FUNCTION StationParameter_28000_1  : BOOL
VAR
  nStationParameter                 : UINT; // THIS IS ONLY FOR EXAMPLE USE, CHECK MAX_STATION MANUALLY
END_VAR

//-----------------------------------------------------------------------------------------------------------------------------------------
//-----------------------------------------------------------------------------------------------------------------------------------------
//
//  HAUD 2026.11.02
//
//  - hard coded station parameters
//  - TODO: xml DataServer implementation for station parameter read/write
//
//  - reminder: (this you HAVE to check manually when setting up the transport)
//-----------------------------------------------------------------------------
//    - DO NOT place the modulo turn within the range of a station
//
//    - in case the extern process requires multiple xts stations, 
//      - the range must be closed and in strict order
//-----------------------------------------------------------------------------------------------------------------------------------------
//-----------------------------------------------------------------------------------------------------------------------------------------
GVL_XTS.StationStartIndex                                         := 142;
GVL_XTS.StationStart.rPosWait                                     :=    5000.0; // for every TRANSPORT_START this physical position may differ from the rPosWait of StationStartIndex station

GVL_XTS.StationStart.rGap                                         :=     110.0;
GVL_XTS.StationStart.rVelo                                        :=   1_250.0;
GVL_XTS.StationStart.rAccDec                                      :=  12_500.0;
GVL_XTS.StationStart.rJerk                                        := 100_000.0;

FOR nStationParameter := 1 TO GVL_XTS_CONSTANTS.MAX_STATION
DO
  GVL_XTS.StationParameter[nStationParameter].eType               := E_STATION_TYPE.STATION_PROCESS;
  GVL_XTS.StationParameter[nStationParameter].rGap                := MAIN_APP.rDefaultGap;
  GVL_XTS.StationParameter[nStationParameter].rVelo               := MAIN_APP.rDefaultVeloMin;
  GVL_XTS.StationParameter[nStationParameter].rAccDec             := MAIN_APP.rDefaultAccDec;
  GVL_XTS.StationParameter[nStationParameter].rJerk               := MAIN_APP.rDefaultJerk;
END_FOR
//-----------------------------------------------------------------------------------------------------------------------------------------
//  PRC 01 reserve
//-----------------------------------------------------------------------------------------------------------------------------------------
FOR nStationParameter := 1 TO 16
DO
  GVL_XTS.StationParameter[nStationParameter].rVelo               := MAIN_APP.rDefaultVeloMin;
END_FOR
nStationParameter := 1;
GVL_XTS.StationParameter[nStationParameter].eType                 := E_STATION_TYPE.STATION_PROCESS;
GVL_XTS.StationParameter[nStationParameter].sText                 := 'PRC_01_01';
GVL_XTS.StationParameter[nStationParameter].nConfiguredStopCount  :=       1;   // how many stops the mover has to make in this station

GVL_XTS.StationParameter[nStationParameter].rPosWait              :=   3000.0+80.0; // absolute modulo position
GVL_XTS.StationParameter[nStationParameter].rPosStop[1]           :=       0.0; // relative to rPosWait
GVL_XTS.StationParameter[nStationParameter].rReleaseDistance      :=    2000.0; // relative to Mover.ActPos

nStationParameter := 2;
GVL_XTS.StationParameter[nStationParameter].eType                 := E_STATION_TYPE.STATION_PROCESS;
GVL_XTS.StationParameter[nStationParameter].sText                 := 'PRC_01_02';
GVL_XTS.StationParameter[nStationParameter].nConfiguredStopCount  :=       1;   // how many stops the mover has to make in this station

GVL_XTS.StationParameter[nStationParameter].rPosWait              :=   3000.0+160.0; // absolute modulo position
GVL_XTS.StationParameter[nStationParameter].rPosStop[1]           :=       0.0; // relative to rPosWait
GVL_XTS.StationParameter[nStationParameter].rReleaseDistance      :=    1900.0; // relative to Mover.ActPos

nStationParameter := 3;
GVL_XTS.StationParameter[nStationParameter].eType                 := E_STATION_TYPE.STATION_PROCESS;
GVL_XTS.StationParameter[nStationParameter].sText                 := 'PRC_01_03';
GVL_XTS.StationParameter[nStationParameter].nConfiguredStopCount  :=       1;   // how many stops the mover has to make in this station

GVL_XTS.StationParameter[nStationParameter].rPosWait              :=     3000.0+240.0; // absolute modulo position
GVL_XTS.StationParameter[nStationParameter].rPosStop[1]           :=       0.0; // relative to rPosWait
GVL_XTS.StationParameter[nStationParameter].rReleaseDistance      :=    1120.0; // relative to Mover.ActPos

nStationParameter := 4;
GVL_XTS.StationParameter[nStationParameter].eType                 := E_STATION_TYPE.STATION_PROCESS;
GVL_XTS.StationParameter[nStationParameter].sText                 := 'PRC_01_04';
GVL_XTS.StationParameter[nStationParameter].nConfiguredStopCount  :=       1;   // how many stops the mover has to make in this station

GVL_XTS.StationParameter[nStationParameter].rPosWait              :=     3000.0+320.0; // absolute modulo position
GVL_XTS.StationParameter[nStationParameter].rPosStop[1]           :=       0.0; // relative to rPosWait
GVL_XTS.StationParameter[nStationParameter].rReleaseDistance      :=    1040.0; // relative to Mover.ActPos

nStationParameter := 5;
GVL_XTS.StationParameter[nStationParameter].eType                 := E_STATION_TYPE.STATION_PROCESS;
GVL_XTS.StationParameter[nStationParameter].sText                 := 'PRC_01_05';
GVL_XTS.StationParameter[nStationParameter].nConfiguredStopCount  :=       1;   // how many stops the mover has to make in this station

GVL_XTS.StationParameter[nStationParameter].rPosWait              :=     3000.0+400.0; // absolute modulo position
GVL_XTS.StationParameter[nStationParameter].rPosStop[1]           :=       0.0; // relative to rPosWait
GVL_XTS.StationParameter[nStationParameter].rReleaseDistance      :=     960.0; // relative to Mover.ActPos

nStationParameter := 6;
GVL_XTS.StationParameter[nStationParameter].eType                 := E_STATION_TYPE.STATION_PROCESS;
GVL_XTS.StationParameter[nStationParameter].sText                 := 'PRC_01_06';
GVL_XTS.StationParameter[nStationParameter].nConfiguredStopCount  :=       1;   // how many stops the mover has to make in this station

GVL_XTS.StationParameter[nStationParameter].rPosWait              :=     3000.0+480.0; // absolute modulo position
GVL_XTS.StationParameter[nStationParameter].rPosStop[1]           :=       0.0; // relative to rPosWait
GVL_XTS.StationParameter[nStationParameter].rReleaseDistance      :=     880.0; // relative to Mover.ActPos

nStationParameter := 7;
GVL_XTS.StationParameter[nStationParameter].eType                 := E_STATION_TYPE.STATION_PROCESS;
GVL_XTS.StationParameter[nStationParameter].sText                 := 'PRC_01_07';
GVL_XTS.StationParameter[nStationParameter].nConfiguredStopCount  :=       1;   // how many stops the mover has to make in this station

GVL_XTS.StationParameter[nStationParameter].rPosWait              :=     3000.0+560.0; // absolute modulo position
GVL_XTS.StationParameter[nStationParameter].rPosStop[1]           :=       0.0; // relative to rPosWait
GVL_XTS.StationParameter[nStationParameter].rReleaseDistance      :=     800.0; // relative to Mover.ActPos

nStationParameter := 8;
GVL_XTS.StationParameter[nStationParameter].eType                 := E_STATION_TYPE.STATION_PROCESS;
GVL_XTS.StationParameter[nStationParameter].sText                 := 'PRC_01_08';
GVL_XTS.StationParameter[nStationParameter].nConfiguredStopCount  :=       1;   // how many stops the mover has to make in this station

GVL_XTS.StationParameter[nStationParameter].rPosWait              :=     3000.0+640.0; // absolute modulo position
GVL_XTS.StationParameter[nStationParameter].rPosStop[1]           :=       0.0; // relative to rPosWait
GVL_XTS.StationParameter[nStationParameter].rReleaseDistance      :=     720.0; // relative to Mover.ActPos

nStationParameter := 9;
GVL_XTS.StationParameter[nStationParameter].eType                 := E_STATION_TYPE.STATION_PROCESS;
GVL_XTS.StationParameter[nStationParameter].sText                 := 'PRC_01_09';
GVL_XTS.StationParameter[nStationParameter].nConfiguredStopCount  :=       1;   // how many stops the mover has to make in this station

GVL_XTS.StationParameter[nStationParameter].rPosWait              :=     3000.0+720.0; // absolute modulo position
GVL_XTS.StationParameter[nStationParameter].rPosStop[1]           :=       0.0; // relative to rPosWait
GVL_XTS.StationParameter[nStationParameter].rReleaseDistance      :=     640.0; // relative to Mover.ActPos

nStationParameter := 10;
GVL_XTS.StationParameter[nStationParameter].eType                 := E_STATION_TYPE.STATION_PROCESS;
GVL_XTS.StationParameter[nStationParameter].sText                 := 'PRC_01_10';
GVL_XTS.StationParameter[nStationParameter].nConfiguredStopCount  :=       1;   // how many stops the mover has to make in this station

GVL_XTS.StationParameter[nStationParameter].rPosWait              :=     3000.0+800; // absolute modulo position
GVL_XTS.StationParameter[nStationParameter].rPosStop[1]           :=       0.0; // relative to rPosWait
GVL_XTS.StationParameter[nStationParameter].rReleaseDistance      :=     560.0; // relative to Mover.ActPos

nStationParameter := 11;
GVL_XTS.StationParameter[nStationParameter].eType                 := E_STATION_TYPE.STATION_PROCESS;
GVL_XTS.StationParameter[nStationParameter].sText                 := 'PRC_01_11';
GVL_XTS.StationParameter[nStationParameter].nConfiguredStopCount  :=       1;   // how many stops the mover has to make in this station

GVL_XTS.StationParameter[nStationParameter].rPosWait              :=     3000.0+880.0; // absolute modulo position
GVL_XTS.StationParameter[nStationParameter].rPosStop[1]           :=       0.0; // relative to rPosWait
GVL_XTS.StationParameter[nStationParameter].rReleaseDistance      :=     480.0; // relative to Mover.ActPos

nStationParameter := 12;
GVL_XTS.StationParameter[nStationParameter].eType                 := E_STATION_TYPE.STATION_PROCESS;
GVL_XTS.StationParameter[nStationParameter].sText                 := 'PRC_01_12';
GVL_XTS.StationParameter[nStationParameter].nConfiguredStopCount  :=       1;   // how many stops the mover has to make in this station

GVL_XTS.StationParameter[nStationParameter].rPosWait              :=     3000.0+960.0; // absolute modulo position
GVL_XTS.StationParameter[nStationParameter].rPosStop[1]           :=       0.0; // relative to rPosWait
GVL_XTS.StationParameter[nStationParameter].rReleaseDistance      :=     400.0; // relative to Mover.ActPos

nStationParameter := 13;
GVL_XTS.StationParameter[nStationParameter].eType                 := E_STATION_TYPE.STATION_PROCESS;
GVL_XTS.StationParameter[nStationParameter].sText                 := 'PRC_01_13';
GVL_XTS.StationParameter[nStationParameter].nConfiguredStopCount  :=       1;   // how many stops the mover has to make in this station

GVL_XTS.StationParameter[nStationParameter].rPosWait              :=     3000.0+1040.0; // absolute modulo position
GVL_XTS.StationParameter[nStationParameter].rPosStop[1]           :=       0.0; // relative to rPosWait
GVL_XTS.StationParameter[nStationParameter].rReleaseDistance      :=     320.0; // relative to Mover.ActPos

nStationParameter := 14;
GVL_XTS.StationParameter[nStationParameter].eType                 := E_STATION_TYPE.STATION_PROCESS;
GVL_XTS.StationParameter[nStationParameter].sText                 := 'PRC_01_14';
GVL_XTS.StationParameter[nStationParameter].nConfiguredStopCount  :=       1;   // how many stops the mover has to make in this station

GVL_XTS.StationParameter[nStationParameter].rPosWait              :=     3000.0+1120.0; // absolute modulo position
GVL_XTS.StationParameter[nStationParameter].rPosStop[1]           :=       0.0; // relative to rPosWait
GVL_XTS.StationParameter[nStationParameter].rReleaseDistance      :=     240.0; // relative to Mover.ActPos

nStationParameter := 15;
GVL_XTS.StationParameter[nStationParameter].eType                 := E_STATION_TYPE.STATION_PROCESS;
GVL_XTS.StationParameter[nStationParameter].sText                 := 'PRC_01_15';
GVL_XTS.StationParameter[nStationParameter].nConfiguredStopCount  :=       1;   // how many stops the mover has to make in this station

GVL_XTS.StationParameter[nStationParameter].rPosWait              :=     3000.0+1200.0; // absolute modulo position
GVL_XTS.StationParameter[nStationParameter].rPosStop[1]           :=       0.0; // relative to rPosWait
GVL_XTS.StationParameter[nStationParameter].rReleaseDistance      :=     160.0; // relative to Mover.ActPos

nStationParameter := 16;
GVL_XTS.StationParameter[nStationParameter].eType                 := E_STATION_TYPE.STATION_PROCESS;
GVL_XTS.StationParameter[nStationParameter].sText                 := 'PRC_01_16';
GVL_XTS.StationParameter[nStationParameter].nConfiguredStopCount  :=       1;   // how many stops the mover has to make in this station

GVL_XTS.StationParameter[nStationParameter].rPosWait              :=     3000.0+1280.0; // absolute modulo position
GVL_XTS.StationParameter[nStationParameter].rPosStop[1]           :=       0.0; // relative to rPosWait
GVL_XTS.StationParameter[nStationParameter].rReleaseDistance      :=      25.0; // relative to Mover.ActPos

//-----------------------------------------------------------------------------------------------------------------------------------------
// PRC 03 Cell loading
//-----------------------------------------------------------------------------------------------------------------------------------------
FOR nStationParameter := 20 TO 35
DO
  GVL_XTS.StationParameter[nStationParameter].rVelo               := 1000.0; //MAIN_APP.rDefaultVeloMin;
END_FOR
nStationParameter := 20;
GVL_XTS.StationParameter[nStationParameter].eType                 := E_STATION_TYPE.STATION_PROCESS;
GVL_XTS.StationParameter[nStationParameter].sText                 := 'PROCESS_INFEED_01';
GVL_XTS.StationParameter[nStationParameter].nConfiguredStopCount  :=       1;   // how many stops the mover has to make in this station

GVL_XTS.StationParameter[nStationParameter].rPosWait              :=    10000.0+80.0; // absolute modulo position
GVL_XTS.StationParameter[nStationParameter].rPosStop[1]           :=       0.0; // relative to rPosWait
GVL_XTS.StationParameter[nStationParameter].rReleaseDistance      :=    1900.0; // relative to Mover.ActPos

nStationParameter := 21;
GVL_XTS.StationParameter[nStationParameter].eType                 := E_STATION_TYPE.STATION_PROCESS;
GVL_XTS.StationParameter[nStationParameter].sText                 := 'PROCESS_INFEED_02';
GVL_XTS.StationParameter[nStationParameter].nConfiguredStopCount  :=       1;   // how many stops the mover has to make in this station

GVL_XTS.StationParameter[nStationParameter].rPosWait              :=    10000.0+160.0; // absolute modulo position
GVL_XTS.StationParameter[nStationParameter].rPosStop[1]           :=       0.0; // relative to rPosWait
GVL_XTS.StationParameter[nStationParameter].rReleaseDistance      :=    1800.0; // relative to Mover.ActPos

nStationParameter := 22;
GVL_XTS.StationParameter[nStationParameter].eType                 := E_STATION_TYPE.STATION_PROCESS;
GVL_XTS.StationParameter[nStationParameter].sText                 := 'PROCESS_INFEED_03';
GVL_XTS.StationParameter[nStationParameter].nConfiguredStopCount  :=       1;   // how many stops the mover has to make in this station

GVL_XTS.StationParameter[nStationParameter].rPosWait              :=    10000.0+240.0; // absolute modulo position
GVL_XTS.StationParameter[nStationParameter].rPosStop[1]           :=       0.0; // relative to rPosWait
GVL_XTS.StationParameter[nStationParameter].rReleaseDistance      :=     1700.0; // relative to Mover.ActPos

nStationParameter := 23;
GVL_XTS.StationParameter[nStationParameter].eType                 := E_STATION_TYPE.STATION_PROCESS;
GVL_XTS.StationParameter[nStationParameter].sText                 := 'PROCESS_INFEED_04';
GVL_XTS.StationParameter[nStationParameter].nConfiguredStopCount  :=       1;   // how many stops the mover has to make in this station

GVL_XTS.StationParameter[nStationParameter].rPosWait              :=    10000.0+320.0; // absolute modulo position
GVL_XTS.StationParameter[nStationParameter].rPosStop[1]           :=       0.0; // relative to rPosWait
GVL_XTS.StationParameter[nStationParameter].rReleaseDistance      :=     1600.0; // relative to Mover.ActPos

nStationParameter := 24;
GVL_XTS.StationParameter[nStationParameter].eType                 := E_STATION_TYPE.STATION_PROCESS;
GVL_XTS.StationParameter[nStationParameter].sText                 := 'PROCESS_INFEED_05';
GVL_XTS.StationParameter[nStationParameter].nConfiguredStopCount  :=       1;   // how many stops the mover has to make in this station

GVL_XTS.StationParameter[nStationParameter].rPosWait              :=    10000.0+400.0; // absolute modulo position
GVL_XTS.StationParameter[nStationParameter].rPosStop[1]           :=       0.0; // relative to rPosWait
GVL_XTS.StationParameter[nStationParameter].rReleaseDistance      :=     1500.0; // relative to Mover.ActPos

nStationParameter := 25;
GVL_XTS.StationParameter[nStationParameter].eType                 := E_STATION_TYPE.STATION_PROCESS;
GVL_XTS.StationParameter[nStationParameter].sText                 := 'PROCESS_INFEED_06';
GVL_XTS.StationParameter[nStationParameter].nConfiguredStopCount  :=       1;   // how many stops the mover has to make in this station

GVL_XTS.StationParameter[nStationParameter].rPosWait              :=    10000.0+480.0; // absolute modulo position
GVL_XTS.StationParameter[nStationParameter].rPosStop[1]           :=       0.0; // relative to rPosWait
GVL_XTS.StationParameter[nStationParameter].rReleaseDistance      :=     1400.0; // relative to Mover.ActPos

nStationParameter := 26;
GVL_XTS.StationParameter[nStationParameter].eType                 := E_STATION_TYPE.STATION_PROCESS;
GVL_XTS.StationParameter[nStationParameter].sText                 := 'PROCESS_INFEED_07';
GVL_XTS.StationParameter[nStationParameter].nConfiguredStopCount  :=       1;   // how many stops the mover has to make in this station

GVL_XTS.StationParameter[nStationParameter].rPosWait              :=    10000.0+560.0; // absolute modulo position
GVL_XTS.StationParameter[nStationParameter].rPosStop[1]           :=       0.0; // relative to rPosWait
GVL_XTS.StationParameter[nStationParameter].rReleaseDistance      :=     640.0; // relative to Mover.ActPos

nStationParameter := 27;
GVL_XTS.StationParameter[nStationParameter].eType                 := E_STATION_TYPE.STATION_PROCESS;
GVL_XTS.StationParameter[nStationParameter].sText                 := 'PROCESS_INFEED_08';
GVL_XTS.StationParameter[nStationParameter].nConfiguredStopCount  :=       1;   // how many stops the mover has to make in this station

GVL_XTS.StationParameter[nStationParameter].rPosWait              :=    10000.0+640.0; // absolute modulo position
GVL_XTS.StationParameter[nStationParameter].rPosStop[1]           :=       0.0; // relative to rPosWait
GVL_XTS.StationParameter[nStationParameter].rReleaseDistance      :=     560.0; // relative to Mover.ActPos

nStationParameter := 28;
GVL_XTS.StationParameter[nStationParameter].eType                 := E_STATION_TYPE.STATION_PROCESS;
GVL_XTS.StationParameter[nStationParameter].sText                 := 'PROCESS_INFEED_09';
GVL_XTS.StationParameter[nStationParameter].nConfiguredStopCount  :=       1;   // how many stops the mover has to make in this station

GVL_XTS.StationParameter[nStationParameter].rPosWait              :=    10000.0+720.0; // absolute modulo position
GVL_XTS.StationParameter[nStationParameter].rPosStop[1]           :=       0.0; // relative to rPosWait
GVL_XTS.StationParameter[nStationParameter].rReleaseDistance      :=     480.0; // relative to Mover.ActPos

nStationParameter := 29;
GVL_XTS.StationParameter[nStationParameter].eType                 := E_STATION_TYPE.STATION_PROCESS;
GVL_XTS.StationParameter[nStationParameter].sText                 := 'PROCESS_INFEED_10';
GVL_XTS.StationParameter[nStationParameter].nConfiguredStopCount  :=       1;   // how many stops the mover has to make in this station

GVL_XTS.StationParameter[nStationParameter].rPosWait              :=    10000.0+800.0; // absolute modulo position
GVL_XTS.StationParameter[nStationParameter].rPosStop[1]           :=       0.0; // relative to rPosWait
GVL_XTS.StationParameter[nStationParameter].rReleaseDistance      :=     400.0; // relative to Mover.ActPos

nStationParameter := 30;
GVL_XTS.StationParameter[nStationParameter].eType                 := E_STATION_TYPE.STATION_PROCESS;
GVL_XTS.StationParameter[nStationParameter].sText                 := 'PROCESS_INFEED_11';
GVL_XTS.StationParameter[nStationParameter].nConfiguredStopCount  :=       1;   // how many stops the mover has to make in this station

GVL_XTS.StationParameter[nStationParameter].rPosWait              :=    10000.0+880.0; // absolute modulo position
GVL_XTS.StationParameter[nStationParameter].rPosStop[1]           :=       0.0; // relative to rPosWait
GVL_XTS.StationParameter[nStationParameter].rReleaseDistance      :=     320.0; // relative to Mover.ActPos

nStationParameter := 31;
GVL_XTS.StationParameter[nStationParameter].eType                 := E_STATION_TYPE.STATION_PROCESS;
GVL_XTS.StationParameter[nStationParameter].sText                 := 'PROCESS_INFEED_12';
GVL_XTS.StationParameter[nStationParameter].nConfiguredStopCount  :=       1;   // how many stops the mover has to make in this station

GVL_XTS.StationParameter[nStationParameter].rPosWait              :=    10000.0+960.0; // absolute modulo position
GVL_XTS.StationParameter[nStationParameter].rPosStop[1]           :=       0.0; // relative to rPosWait
GVL_XTS.StationParameter[nStationParameter].rReleaseDistance      :=     240.0; // relative to Mover.ActPos

nStationParameter := 32;
GVL_XTS.StationParameter[nStationParameter].eType                 := E_STATION_TYPE.STATION_PROCESS;
GVL_XTS.StationParameter[nStationParameter].sText                 := 'PROCESS_INFEED_13';
GVL_XTS.StationParameter[nStationParameter].nConfiguredStopCount  :=       1;   // how many stops the mover has to make in this station

GVL_XTS.StationParameter[nStationParameter].rPosWait              :=    10000.0+1040.0; // absolute modulo position
GVL_XTS.StationParameter[nStationParameter].rPosStop[1]           :=       0.0; // relative to rPosWait
GVL_XTS.StationParameter[nStationParameter].rReleaseDistance      :=     160.0; // relative to Mover.ActPos

nStationParameter := 33;
GVL_XTS.StationParameter[nStationParameter].eType                 := E_STATION_TYPE.STATION_PROCESS;
GVL_XTS.StationParameter[nStationParameter].sText                 := 'PROCESS_INFEED_14';
GVL_XTS.StationParameter[nStationParameter].nConfiguredStopCount  :=       1;   // how many stops the mover has to make in this station

GVL_XTS.StationParameter[nStationParameter].rPosWait              :=    10000.0+1120.0; // absolute modulo position
GVL_XTS.StationParameter[nStationParameter].rPosStop[1]           :=       0.0; // relative to rPosWait
GVL_XTS.StationParameter[nStationParameter].rReleaseDistance      :=      80.0; // relative to Mover.ActPos

nStationParameter := 34;
GVL_XTS.StationParameter[nStationParameter].eType                 := E_STATION_TYPE.STATION_PROCESS;
GVL_XTS.StationParameter[nStationParameter].sText                 := 'PROCESS_INFEED_15';
GVL_XTS.StationParameter[nStationParameter].nConfiguredStopCount  :=       1;   // how many stops the mover has to make in this station

GVL_XTS.StationParameter[nStationParameter].rPosWait              :=    10000.0+1200.0; // absolute modulo position
GVL_XTS.StationParameter[nStationParameter].rPosStop[1]           :=       0.0; // relative to rPosWait
GVL_XTS.StationParameter[nStationParameter].rReleaseDistance      :=      25.0; // relative to Mover.ActPos

nStationParameter := 35;
GVL_XTS.StationParameter[nStationParameter].eType                 := E_STATION_TYPE.STATION_PROCESS;
GVL_XTS.StationParameter[nStationParameter].sText                 := 'PROCESS_INFEED_16';
GVL_XTS.StationParameter[nStationParameter].nConfiguredStopCount  :=       1;   // how many stops the mover has to make in this station

GVL_XTS.StationParameter[nStationParameter].rPosWait              :=    10000.0+1280.0; // absolute modulo position
GVL_XTS.StationParameter[nStationParameter].rPosStop[1]           :=       0.0; // relative to rPosWait
GVL_XTS.StationParameter[nStationParameter].rReleaseDistance      :=      -5.0; // relative to Mover.ActPos

//-----------------------------------------------------------------------------------------------------------------------------------------
// CONTINUOUS_CLEAN
//-----------------------------------------------------------------------------------------------------------------------------------------
nStationParameter := 37;
GVL_XTS.StationParameter[nStationParameter].eType                 := E_STATION_TYPE.STATION_PROCESS;
GVL_XTS.StationParameter[nStationParameter].sText                 := 'CONTINUOUS_CLEAN';
GVL_XTS.StationParameter[nStationParameter].nConfiguredStopCount  :=       1;   // how many stops the mover has to make in this station

GVL_XTS.StationParameter[nStationParameter].rPosWait              :=   12900.0; // absolute modulo position
GVL_XTS.StationParameter[nStationParameter].rPosStop[1]           :=       0.0; // relative to rPosWait
GVL_XTS.StationParameter[nStationParameter].rReleaseDistance      :=     -10.0; // relative to Mover.ActPos
GVL_XTS.StationParameter[nStationParameter].rVelo                 :=     1100.0;
GVL_XTS.StationParameter[nStationParameter].rGap                  :=     110.0;

//-----------------------------------------------------------------------------------------------------------------------------------------
// CONTINUOUS_SCAN
//-----------------------------------------------------------------------------------------------------------------------------------------
nStationParameter := 38;
GVL_XTS.StationParameter[nStationParameter].eType                 := E_STATION_TYPE.STATION_PROCESS;
GVL_XTS.StationParameter[nStationParameter].sText                 := 'CONTINUOUS_SCAN';
GVL_XTS.StationParameter[nStationParameter].nConfiguredStopCount  :=       1;   // how many stops the mover has to make in this station

GVL_XTS.StationParameter[nStationParameter].rPosWait              :=   14000.0; // absolute modulo position
GVL_XTS.StationParameter[nStationParameter].rPosStop[1]           :=       0.0; // relative to rPosWait
GVL_XTS.StationParameter[nStationParameter].rReleaseDistance      :=     -10.0; // relative to Mover.ActPos
GVL_XTS.StationParameter[nStationParameter].rVelo                 :=     1100.0;
GVL_XTS.StationParameter[nStationParameter].rGap                  :=     110.0;

//-----------------------------------------------------------------------------------------------------------------------------------------
// CONTINUOUS_CAM
//-----------------------------------------------------------------------------------------------------------------------------------------
nStationParameter := 39;
GVL_XTS.StationParameter[nStationParameter].eType                 := E_STATION_TYPE.STATION_PROCESS;
GVL_XTS.StationParameter[nStationParameter].sText                 := 'CONTINUOUS_CAM';
GVL_XTS.StationParameter[nStationParameter].nConfiguredStopCount  :=       1;   // how many stops the mover has to make in this station

GVL_XTS.StationParameter[nStationParameter].rPosWait              :=   14300.0; // absolute modulo position
GVL_XTS.StationParameter[nStationParameter].rPosStop[1]           :=       0.0; // relative to rPosWait
GVL_XTS.StationParameter[nStationParameter].rReleaseDistance      :=     -10.0; // relative to Mover.ActPos
GVL_XTS.StationParameter[nStationParameter].rVelo                 :=     1100.0;
GVL_XTS.StationParameter[nStationParameter].rGap                  :=     109.0;

//-----------------------------------------------------------------------------------------------------------------------------------------
// DISTRIBUTOR_ASSEMBLY_01
//-----------------------------------------------------------------------------------------------------------------------------------------
nStationParameter := 40;
GVL_XTS.StationParameter[nStationParameter].eType                 := E_STATION_TYPE.STATION_PROCESS;
GVL_XTS.StationParameter[nStationParameter].sText                 := 'DISTRIBUTOR_ASSEMBLY_01';
GVL_XTS.StationParameter[nStationParameter].nConfiguredStopCount  :=       1;   // how many stops the mover has to make in this station

GVL_XTS.StationParameter[nStationParameter].rPosWait              :=   15250.0; // absolute modulo position
GVL_XTS.StationParameter[nStationParameter].rPosStop[1]           :=       0.0; // relative to rPosWait
GVL_XTS.StationParameter[nStationParameter].rReleaseDistance      :=     -10.0; // relative to Mover.ActPos
GVL_XTS.StationParameter[nStationParameter].rVelo                 :=    1500.0;
GVL_XTS.StationParameter[nStationParameter].rGap                  :=     109.0;

//-----------------------------------------------------------------------------------------------------------------------------------------
// PRC 05 Visual check film bottom
//-----------------------------------------------------------------------------------------------------------------------------------------
FOR nStationParameter := 41 TO 56
DO
  GVL_XTS.StationParameter[nStationParameter].rVelo               := MAIN_APP.rDefaultVeloMin;
END_FOR
nStationParameter := 41;
GVL_XTS.StationParameter[nStationParameter].eType                 := E_STATION_TYPE.STATION_PROCESS;
GVL_XTS.StationParameter[nStationParameter].sText                 := 'PROCESS_ASSEMBLY_01_01';
GVL_XTS.StationParameter[nStationParameter].nConfiguredStopCount  :=       1;   // how many stops the mover has to make in this station

GVL_XTS.StationParameter[nStationParameter].rPosWait              :=    15500.0+110.0; // absolute modulo position
GVL_XTS.StationParameter[nStationParameter].rPosStop[1]           :=       0.0; // relative to rPosWait
GVL_XTS.StationParameter[nStationParameter].rReleaseDistance      :=    1540.0; // relative to Mover.ActPos
GVL_XTS.StationParameter[nStationParameter].rGap                  :=     109.0;

nStationParameter := 42;
GVL_XTS.StationParameter[nStationParameter].eType                 := E_STATION_TYPE.STATION_PROCESS;
GVL_XTS.StationParameter[nStationParameter].sText                 := 'PROCESS_ASSEMBLY_01_02';
GVL_XTS.StationParameter[nStationParameter].nConfiguredStopCount  :=       1;   // how many stops the mover has to make in this station

GVL_XTS.StationParameter[nStationParameter].rPosWait              :=    15500.0+220.0; // absolute modulo position
GVL_XTS.StationParameter[nStationParameter].rPosStop[1]           :=       0.0; // relative to rPosWait
GVL_XTS.StationParameter[nStationParameter].rReleaseDistance      :=     1430.0; // relative to Mover.ActPos
GVL_XTS.StationParameter[nStationParameter].rGap                  :=     109.0;

nStationParameter := 43;
GVL_XTS.StationParameter[nStationParameter].eType                 := E_STATION_TYPE.STATION_PROCESS;
GVL_XTS.StationParameter[nStationParameter].sText                 := 'PROCESS_ASSEMBLY_01_03';
GVL_XTS.StationParameter[nStationParameter].nConfiguredStopCount  :=       1;   // how many stops the mover has to make in this station

GVL_XTS.StationParameter[nStationParameter].rPosWait              :=    15500.0+330.0; // absolute modulo position
GVL_XTS.StationParameter[nStationParameter].rPosStop[1]           :=       0.0; // relative to rPosWait
GVL_XTS.StationParameter[nStationParameter].rReleaseDistance      :=     1320.0; // relative to Mover.ActPos
GVL_XTS.StationParameter[nStationParameter].rGap                  :=     109.0;

nStationParameter := 44;
GVL_XTS.StationParameter[nStationParameter].eType                 := E_STATION_TYPE.STATION_PROCESS;
GVL_XTS.StationParameter[nStationParameter].sText                 := 'PROCESS_ASSEMBLY_01_04';
GVL_XTS.StationParameter[nStationParameter].nConfiguredStopCount  :=       1;   // how many stops the mover has to make in this station

GVL_XTS.StationParameter[nStationParameter].rPosWait              :=    15500.0+440.0; // absolute modulo position
GVL_XTS.StationParameter[nStationParameter].rPosStop[1]           :=       0.0; // relative to rPosWait
GVL_XTS.StationParameter[nStationParameter].rReleaseDistance      :=     1210.0; // relative to Mover.ActPos
GVL_XTS.StationParameter[nStationParameter].rGap                  :=     109.0;

nStationParameter := 45;
GVL_XTS.StationParameter[nStationParameter].eType                 := E_STATION_TYPE.STATION_PROCESS;
GVL_XTS.StationParameter[nStationParameter].sText                 := 'PROCESS_ASSEMBLY_01_05';
GVL_XTS.StationParameter[nStationParameter].nConfiguredStopCount  :=       1;   // how many stops the mover has to make in this station

GVL_XTS.StationParameter[nStationParameter].rPosWait              :=    15500.0+550.0; // absolute modulo position
GVL_XTS.StationParameter[nStationParameter].rPosStop[1]           :=       0.0; // relative to rPosWait
GVL_XTS.StationParameter[nStationParameter].rReleaseDistance      :=     1100.0; // relative to Mover.ActPos
GVL_XTS.StationParameter[nStationParameter].rGap                  :=     109.0;

nStationParameter := 46;
GVL_XTS.StationParameter[nStationParameter].eType                 := E_STATION_TYPE.STATION_PROCESS;
GVL_XTS.StationParameter[nStationParameter].sText                 := 'PROCESS_ASSEMBLY_01_06';
GVL_XTS.StationParameter[nStationParameter].nConfiguredStopCount  :=       1;   // how many stops the mover has to make in this station

GVL_XTS.StationParameter[nStationParameter].rPosWait              :=    15500.0+660.0; // absolute modulo position
GVL_XTS.StationParameter[nStationParameter].rPosStop[1]           :=       0.0; // relative to rPosWait
GVL_XTS.StationParameter[nStationParameter].rReleaseDistance      :=     990.0; // relative to Mover.ActPos
GVL_XTS.StationParameter[nStationParameter].rGap                  :=     109.0;

nStationParameter := 47;
GVL_XTS.StationParameter[nStationParameter].eType                 := E_STATION_TYPE.STATION_PROCESS;
GVL_XTS.StationParameter[nStationParameter].sText                 := 'PROCESS_ASSEMBLY_01_07';
GVL_XTS.StationParameter[nStationParameter].nConfiguredStopCount  :=       1;   // how many stops the mover has to make in this station

GVL_XTS.StationParameter[nStationParameter].rPosWait              :=    15500.0+770.0; // absolute modulo position
GVL_XTS.StationParameter[nStationParameter].rPosStop[1]           :=       0.0; // relative to rPosWait
GVL_XTS.StationParameter[nStationParameter].rReleaseDistance      :=     880.0; // relative to Mover.ActPos
GVL_XTS.StationParameter[nStationParameter].rGap                  :=     109.0;

nStationParameter := 48;
GVL_XTS.StationParameter[nStationParameter].eType                 := E_STATION_TYPE.STATION_PROCESS;
GVL_XTS.StationParameter[nStationParameter].sText                 := 'PROCESS_ASSEMBLY_01_08';
GVL_XTS.StationParameter[nStationParameter].nConfiguredStopCount  :=       1;   // how many stops the mover has to make in this station

GVL_XTS.StationParameter[nStationParameter].rPosWait              :=    15500.0+880.0; // absolute modulo position
GVL_XTS.StationParameter[nStationParameter].rPosStop[1]           :=       0.0; // relative to rPosWait
GVL_XTS.StationParameter[nStationParameter].rReleaseDistance      :=     770.0; // relative to Mover.ActPos
GVL_XTS.StationParameter[nStationParameter].rGap                  :=     109.0;

nStationParameter := 49;
GVL_XTS.StationParameter[nStationParameter].eType                 := E_STATION_TYPE.STATION_PROCESS;
GVL_XTS.StationParameter[nStationParameter].sText                 := 'PROCESS_ASSEMBLY_01_09';
GVL_XTS.StationParameter[nStationParameter].nConfiguredStopCount  :=       1;   // how many stops the mover has to make in this station

GVL_XTS.StationParameter[nStationParameter].rPosWait              :=    15500.0+990.0; // absolute modulo position
GVL_XTS.StationParameter[nStationParameter].rPosStop[1]           :=       0.0; // relative to rPosWait
GVL_XTS.StationParameter[nStationParameter].rReleaseDistance      :=     660.0; // relative to Mover.ActPos
GVL_XTS.StationParameter[nStationParameter].rGap                  :=     109.0;

nStationParameter := 50;
GVL_XTS.StationParameter[nStationParameter].eType                 := E_STATION_TYPE.STATION_PROCESS;
GVL_XTS.StationParameter[nStationParameter].sText                 := 'PROCESS_ASSEMBLY_01_10';
GVL_XTS.StationParameter[nStationParameter].nConfiguredStopCount  :=       1;   // how many stops the mover has to make in this station

GVL_XTS.StationParameter[nStationParameter].rPosWait              :=    15500.0+1100.0; // absolute modulo position
GVL_XTS.StationParameter[nStationParameter].rPosStop[1]           :=       0.0; // relative to rPosWait
GVL_XTS.StationParameter[nStationParameter].rReleaseDistance      :=     550.0; // relative to Mover.ActPos
GVL_XTS.StationParameter[nStationParameter].rGap                  :=     109.0;

nStationParameter := 51;
GVL_XTS.StationParameter[nStationParameter].eType                 := E_STATION_TYPE.STATION_PROCESS;
GVL_XTS.StationParameter[nStationParameter].sText                 := 'PROCESS_ASSEMBLY_01_11';
GVL_XTS.StationParameter[nStationParameter].nConfiguredStopCount  :=       1;   // how many stops the mover has to make in this station

GVL_XTS.StationParameter[nStationParameter].rPosWait              :=    15500.0+1210.0; // absolute modulo position
GVL_XTS.StationParameter[nStationParameter].rPosStop[1]           :=       0.0; // relative to rPosWait
GVL_XTS.StationParameter[nStationParameter].rReleaseDistance      :=     440.0; // relative to Mover.ActPos
GVL_XTS.StationParameter[nStationParameter].rGap                  :=     109.0;

nStationParameter := 52;
GVL_XTS.StationParameter[nStationParameter].eType                 := E_STATION_TYPE.STATION_PROCESS;
GVL_XTS.StationParameter[nStationParameter].sText                 := 'PROCESS_ASSEMBLY_01_12';
GVL_XTS.StationParameter[nStationParameter].nConfiguredStopCount  :=       1;   // how many stops the mover has to make in this station

GVL_XTS.StationParameter[nStationParameter].rPosWait              :=    15500.0+1320.0; // absolute modulo position
GVL_XTS.StationParameter[nStationParameter].rPosStop[1]           :=       0.0; // relative to rPosWait
GVL_XTS.StationParameter[nStationParameter].rReleaseDistance      :=     330.0; // relative to Mover.ActPos
GVL_XTS.StationParameter[nStationParameter].rGap                  :=     109.0;

nStationParameter := 53;
GVL_XTS.StationParameter[nStationParameter].eType                 := E_STATION_TYPE.STATION_PROCESS;
GVL_XTS.StationParameter[nStationParameter].sText                 := 'PROCESS_ASSEMBLY_01_13';
GVL_XTS.StationParameter[nStationParameter].nConfiguredStopCount  :=       1;   // how many stops the mover has to make in this station

GVL_XTS.StationParameter[nStationParameter].rPosWait              :=    15500.0+1430.0; // absolute modulo position
GVL_XTS.StationParameter[nStationParameter].rPosStop[1]           :=       0.0; // relative to rPosWait
GVL_XTS.StationParameter[nStationParameter].rReleaseDistance      :=     220.0; // relative to Mover.ActPos
GVL_XTS.StationParameter[nStationParameter].rGap                  :=     109.0;

nStationParameter := 54;
GVL_XTS.StationParameter[nStationParameter].eType                 := E_STATION_TYPE.STATION_PROCESS;
GVL_XTS.StationParameter[nStationParameter].sText                 := 'PROCESS_ASSEMBLY_01_14';
GVL_XTS.StationParameter[nStationParameter].nConfiguredStopCount  :=       1;   // how many stops the mover has to make in this station

GVL_XTS.StationParameter[nStationParameter].rPosWait              :=    15500.0+1540.0; // absolute modulo position
GVL_XTS.StationParameter[nStationParameter].rPosStop[1]           :=       0.0; // relative to rPosWait
GVL_XTS.StationParameter[nStationParameter].rReleaseDistance      :=     110.0; // relative to Mover.ActPos
GVL_XTS.StationParameter[nStationParameter].rGap                  :=     109.0;

nStationParameter := 55;
GVL_XTS.StationParameter[nStationParameter].eType                 := E_STATION_TYPE.STATION_PROCESS;
GVL_XTS.StationParameter[nStationParameter].sText                 := 'PROCESS_ASSEMBLY_01_15';
GVL_XTS.StationParameter[nStationParameter].nConfiguredStopCount  :=       1;   // how many stops the mover has to make in this station

GVL_XTS.StationParameter[nStationParameter].rPosWait              :=    15500.0+1650.0; // absolute modulo position
GVL_XTS.StationParameter[nStationParameter].rPosStop[1]           :=       0.0; // relative to rPosWait
GVL_XTS.StationParameter[nStationParameter].rReleaseDistance      :=      25.0; // relative to Mover.ActPos
GVL_XTS.StationParameter[nStationParameter].rGap                  :=     109.0;

nStationParameter := 56;
GVL_XTS.StationParameter[nStationParameter].eType                 := E_STATION_TYPE.STATION_PROCESS;
GVL_XTS.StationParameter[nStationParameter].sText                 := 'PROCESS_ASSEMBLY_01_16';
GVL_XTS.StationParameter[nStationParameter].nConfiguredStopCount  :=       1;   // how many stops the mover has to make in this station

GVL_XTS.StationParameter[nStationParameter].rPosWait              :=    15500.0+1760.0; // absolute modulo position
GVL_XTS.StationParameter[nStationParameter].rPosStop[1]           :=       0.0; // relative to rPosWait
GVL_XTS.StationParameter[nStationParameter].rReleaseDistance      :=      -5.0; // relative to Mover.ActPos
GVL_XTS.StationParameter[nStationParameter].rGap                  :=     109.0;
//-----------------------------------------------------------------------------------------------------------------------------------------
// DISTRIBUTOR_ASSEMBLY_02
//-----------------------------------------------------------------------------------------------------------------------------------------
nStationParameter := 57;
GVL_XTS.StationParameter[nStationParameter].eType                 := E_STATION_TYPE.STATION_PROCESS;
GVL_XTS.StationParameter[nStationParameter].sText                 := 'DISTRIBUTOR_ASSEMBLY_02';
GVL_XTS.StationParameter[nStationParameter].nConfiguredStopCount  :=       1;   // how many stops the mover has to make in this station

GVL_XTS.StationParameter[nStationParameter].rPosWait              :=   18000.0; // absolute modulo position
GVL_XTS.StationParameter[nStationParameter].rPosStop[1]           :=       0.0; // relative to rPosWait
GVL_XTS.StationParameter[nStationParameter].rReleaseDistance      :=      -5.0; // relative to Mover.ActPos
GVL_XTS.StationParameter[nStationParameter].rVelo                 := MAIN_APP.rDefaultVeloMin;

//-----------------------------------------------------------------------------------------------------------------------------------------
// PROCESS_ASSEMBLY_02
//-----------------------------------------------------------------------------------------------------------------------------------------
FOR nStationParameter := 58 TO 69
DO
   GVL_XTS.StationParameter[nStationParameter].rVelo               := MAIN_APP.rDefaultVeloMin;
END_FOR
nStationParameter := 58;
GVL_XTS.StationParameter[nStationParameter].eType                 := E_STATION_TYPE.STATION_PROCESS;
GVL_XTS.StationParameter[nStationParameter].sText                 := 'PROCESS_ASSEMBLY_02_01';
GVL_XTS.StationParameter[nStationParameter].nConfiguredStopCount  :=       1;   // how many stops the mover has to make in this station

GVL_XTS.StationParameter[nStationParameter].rPosWait              :=    19500.0+80.0; // absolute modulo position
GVL_XTS.StationParameter[nStationParameter].rPosStop[1]           :=       0.0; // relative to rPosWait
GVL_XTS.StationParameter[nStationParameter].rReleaseDistance      :=     640.0; // relative to Mover.ActPos

nStationParameter := 59;
GVL_XTS.StationParameter[nStationParameter].eType                 := E_STATION_TYPE.STATION_PROCESS;
GVL_XTS.StationParameter[nStationParameter].sText                 := 'PROCESS_ASSEMBLY_02_02';
GVL_XTS.StationParameter[nStationParameter].nConfiguredStopCount  :=       1;   // how many stops the mover has to make in this station

GVL_XTS.StationParameter[nStationParameter].rPosWait              :=    19500.0+160.0; // absolute modulo position
GVL_XTS.StationParameter[nStationParameter].rPosStop[1]           :=       0.0; // relative to rPosWait
GVL_XTS.StationParameter[nStationParameter].rReleaseDistance      :=     560.0; // relative to Mover.ActPos

nStationParameter := 60;
GVL_XTS.StationParameter[nStationParameter].eType                 := E_STATION_TYPE.STATION_PROCESS;
GVL_XTS.StationParameter[nStationParameter].sText                 := 'PROCESS_ASSEMBLY_02_03';
GVL_XTS.StationParameter[nStationParameter].nConfiguredStopCount  :=       1;   // how many stops the mover has to make in this station

GVL_XTS.StationParameter[nStationParameter].rPosWait              :=    19500.0+240.0; // absolute modulo position
GVL_XTS.StationParameter[nStationParameter].rPosStop[1]           :=       0.0; // relative to rPosWait
GVL_XTS.StationParameter[nStationParameter].rReleaseDistance      :=     480.0; // relative to Mover.ActPos

nStationParameter := 61;
GVL_XTS.StationParameter[nStationParameter].eType                 := E_STATION_TYPE.STATION_PROCESS;
GVL_XTS.StationParameter[nStationParameter].sText                 := 'PROCESS_ASSEMBLY_02_04';
GVL_XTS.StationParameter[nStationParameter].nConfiguredStopCount  :=       1;   // how many stops the mover has to make in this station

GVL_XTS.StationParameter[nStationParameter].rPosWait              :=    19500.0+320.0; // absolute modulo position
GVL_XTS.StationParameter[nStationParameter].rPosStop[1]           :=       0.0; // relative to rPosWait
GVL_XTS.StationParameter[nStationParameter].rReleaseDistance      :=     400.0; // relative to Mover.ActPos

nStationParameter := 62;
GVL_XTS.StationParameter[nStationParameter].eType                 := E_STATION_TYPE.STATION_PROCESS;
GVL_XTS.StationParameter[nStationParameter].sText                 := 'PROCESS_ASSEMBLY_02_05';
GVL_XTS.StationParameter[nStationParameter].nConfiguredStopCount  :=       1;   // how many stops the mover has to make in this station

GVL_XTS.StationParameter[nStationParameter].rPosWait              :=    19500.0+400.0; // absolute modulo position
GVL_XTS.StationParameter[nStationParameter].rPosStop[1]           :=       0.0; // relative to rPosWait
GVL_XTS.StationParameter[nStationParameter].rReleaseDistance      :=      320.0; // relative to Mover.ActPos

nStationParameter := 63;
GVL_XTS.StationParameter[nStationParameter].eType                 := E_STATION_TYPE.STATION_PROCESS;
GVL_XTS.StationParameter[nStationParameter].sText                 := 'PROCESS_ASSEMBLY_02_06';
GVL_XTS.StationParameter[nStationParameter].nConfiguredStopCount  :=       1;   // how many stops the mover has to make in this station

GVL_XTS.StationParameter[nStationParameter].rPosWait              :=    19500.0+480.0; // absolute modulo position
GVL_XTS.StationParameter[nStationParameter].rPosStop[1]           :=       0.0; // relative to rPosWait
GVL_XTS.StationParameter[nStationParameter].rReleaseDistance      :=      240.0; // relative to Mover.ActPos

nStationParameter := 64;
GVL_XTS.StationParameter[nStationParameter].eType                 := E_STATION_TYPE.STATION_PROCESS;
GVL_XTS.StationParameter[nStationParameter].sText                 := 'PROCESS_ASSEMBLY_02_07';
GVL_XTS.StationParameter[nStationParameter].nConfiguredStopCount  :=       1;   // how many stops the mover has to make in this station

GVL_XTS.StationParameter[nStationParameter].rPosWait              :=    19500.0+560.0; // absolute modulo position
GVL_XTS.StationParameter[nStationParameter].rPosStop[1]           :=       0.0; // relative to rPosWait
GVL_XTS.StationParameter[nStationParameter].rReleaseDistance      :=      160.0; // relative to Mover.ActPos

nStationParameter := 65;
GVL_XTS.StationParameter[nStationParameter].eType                 := E_STATION_TYPE.STATION_PROCESS;
GVL_XTS.StationParameter[nStationParameter].sText                 := 'PROCESS_ASSEMBLY_02_08';
GVL_XTS.StationParameter[nStationParameter].nConfiguredStopCount  :=       1;   // how many stops the mover has to make in this station

GVL_XTS.StationParameter[nStationParameter].rPosWait              :=    19500.0+640.0; // absolute modulo position
GVL_XTS.StationParameter[nStationParameter].rPosStop[1]           :=       0.0; // relative to rPosWait
GVL_XTS.StationParameter[nStationParameter].rReleaseDistance      :=     80.0; // relative to Mover.ActPos

nStationParameter := 66;
GVL_XTS.StationParameter[nStationParameter].eType                 := E_STATION_TYPE.STATION_PROCESS;
GVL_XTS.StationParameter[nStationParameter].sText                 := 'PROCESS_ASSEMBLY_02_09';
GVL_XTS.StationParameter[nStationParameter].nConfiguredStopCount  :=       1;   // how many stops the mover has to make in this station

GVL_XTS.StationParameter[nStationParameter].rPosWait              :=    19500.0+720.0; // absolute modulo position
GVL_XTS.StationParameter[nStationParameter].rPosStop[1]           :=       0.0; // relative to rPosWait
GVL_XTS.StationParameter[nStationParameter].rReleaseDistance      :=     25.0; // relative to Mover.ActPos

nStationParameter := 67;
GVL_XTS.StationParameter[nStationParameter].eType                 := E_STATION_TYPE.STATION_PROCESS;
GVL_XTS.StationParameter[nStationParameter].sText                 := 'PROCESS_ASSEMBLY_02_10';
GVL_XTS.StationParameter[nStationParameter].nConfiguredStopCount  :=       1;   // how many stops the mover has to make in this station

GVL_XTS.StationParameter[nStationParameter].rPosWait              :=    19500.0+800.0; // absolute modulo position
GVL_XTS.StationParameter[nStationParameter].rPosStop[1]           :=       0.0; // relative to rPosWait
GVL_XTS.StationParameter[nStationParameter].rReleaseDistance      :=     -5.0; // relative to Mover.ActPos

nStationParameter := 68;
GVL_XTS.StationParameter[nStationParameter].eType                 := E_STATION_TYPE.STATION_PROCESS;
GVL_XTS.StationParameter[nStationParameter].sText                 := 'PROCESS_ASSEMBLY_02_11';
GVL_XTS.StationParameter[nStationParameter].nConfiguredStopCount  :=       1;   // how many stops the mover has to make in this station

GVL_XTS.StationParameter[nStationParameter].rPosWait              :=    19500.0+880.0; // absolute modulo position
GVL_XTS.StationParameter[nStationParameter].rPosStop[1]           :=       0.0; // relative to rPosWait
GVL_XTS.StationParameter[nStationParameter].rReleaseDistance      :=      80.0; // relative to Mover.ActPos

nStationParameter := 69;
GVL_XTS.StationParameter[nStationParameter].eType                 := E_STATION_TYPE.STATION_PROCESS;
GVL_XTS.StationParameter[nStationParameter].sText                 := 'PROCESS_ASSEMBLY_02_12';
GVL_XTS.StationParameter[nStationParameter].nConfiguredStopCount  :=       1;   // how many stops the mover has to make in this station

GVL_XTS.StationParameter[nStationParameter].rPosWait              :=    19500.0+960.0; // absolute modulo position
GVL_XTS.StationParameter[nStationParameter].rPosStop[1]           :=       0.0; // relative to rPosWait
GVL_XTS.StationParameter[nStationParameter].rReleaseDistance      :=      25.0; // relative to Mover.ActPos

//-----------------------------------------------------------------------------------------------------------------------------------------
// DISTRIBUTOR_ASSEMBLY_TEST
//-----------------------------------------------------------------------------------------------------------------------------------------
nStationParameter := 70;
GVL_XTS.StationParameter[nStationParameter].eType                 := E_STATION_TYPE.STATION_PROCESS;
GVL_XTS.StationParameter[nStationParameter].sText                 := 'DISTRIBUTOR_ASSEMBLY_TEST';
GVL_XTS.StationParameter[nStationParameter].nConfiguredStopCount  :=       1;   // how many stops the mover has to make in this station

GVL_XTS.StationParameter[nStationParameter].rPosWait              :=   21000.0; // absolute modulo position
GVL_XTS.StationParameter[nStationParameter].rPosStop[1]           :=       0.0; // relative to rPosWait
GVL_XTS.StationParameter[nStationParameter].rReleaseDistance      :=      -5.0; // relative to Mover.ActPos


//-----------------------------------------------------------------------------------------------------------------------------------------
// PROCESS_ASSEMBLY_TEST
//-----------------------------------------------------------------------------------------------------------------------------------------
FOR nStationParameter := 71 TO 86
DO
   GVL_XTS.StationParameter[nStationParameter].rVelo               := 1000.0;//MAIN_APP.rDefaultVeloMin;
END_FOR
nStationParameter := 71;
GVL_XTS.StationParameter[nStationParameter].eType                 := E_STATION_TYPE.STATION_PROCESS;
GVL_XTS.StationParameter[nStationParameter].sText                 := 'PROCESS_ASSEMBLY_TEST_01';
GVL_XTS.StationParameter[nStationParameter].nConfiguredStopCount  :=       1;   // how many stops the mover has to make in this station

GVL_XTS.StationParameter[nStationParameter].rPosWait              :=    21500.0+80.0; // absolute modulo position
GVL_XTS.StationParameter[nStationParameter].rPosStop[1]           :=       0.0; // relative to rPosWait
GVL_XTS.StationParameter[nStationParameter].rReleaseDistance      :=     1120.0; // relative to Mover.ActPos

nStationParameter := 72;
GVL_XTS.StationParameter[nStationParameter].eType                 := E_STATION_TYPE.STATION_PROCESS;
GVL_XTS.StationParameter[nStationParameter].sText                 := 'PROCESS_ASSEMBLY_TEST_02';
GVL_XTS.StationParameter[nStationParameter].nConfiguredStopCount  :=       1;   // how many stops the mover has to make in this station

GVL_XTS.StationParameter[nStationParameter].rPosWait              :=    21500.0+160.0; // absolute modulo position
GVL_XTS.StationParameter[nStationParameter].rPosStop[1]           :=       0.0; // relative to rPosWait
GVL_XTS.StationParameter[nStationParameter].rReleaseDistance      :=     1040.0; // relative to Mover.ActPos

nStationParameter := 73;
GVL_XTS.StationParameter[nStationParameter].eType                 := E_STATION_TYPE.STATION_PROCESS;
GVL_XTS.StationParameter[nStationParameter].sText                 := 'PROCESS_ASSEMBLY_TEST_03';
GVL_XTS.StationParameter[nStationParameter].nConfiguredStopCount  :=       1;   // how many stops the mover has to make in this station

GVL_XTS.StationParameter[nStationParameter].rPosWait              :=    21500.0+240.0; // absolute modulo position
GVL_XTS.StationParameter[nStationParameter].rPosStop[1]           :=       0.0; // relative to rPosWait
GVL_XTS.StationParameter[nStationParameter].rReleaseDistance      :=    960.0; // relative to Mover.ActPos

nStationParameter := 74;
GVL_XTS.StationParameter[nStationParameter].eType                 := E_STATION_TYPE.STATION_PROCESS;
GVL_XTS.StationParameter[nStationParameter].sText                 := 'PROCESS_ASSEMBLY_TEST_04';
GVL_XTS.StationParameter[nStationParameter].nConfiguredStopCount  :=       1;   // how many stops the mover has to make in this station

GVL_XTS.StationParameter[nStationParameter].rPosWait              :=    21500.0+320.0; // absolute modulo position
GVL_XTS.StationParameter[nStationParameter].rPosStop[1]           :=       0.0; // relative to rPosWait
GVL_XTS.StationParameter[nStationParameter].rReleaseDistance      :=     880.0; // relative to Mover.ActPos

nStationParameter := 75;
GVL_XTS.StationParameter[nStationParameter].eType                 := E_STATION_TYPE.STATION_PROCESS;
GVL_XTS.StationParameter[nStationParameter].sText                 := 'PROCESS_ASSEMBLY_TEST_05';
GVL_XTS.StationParameter[nStationParameter].nConfiguredStopCount  :=       1;   // how many stops the mover has to make in this station

GVL_XTS.StationParameter[nStationParameter].rPosWait              :=    21500.0+400.0; // absolute modulo position
GVL_XTS.StationParameter[nStationParameter].rPosStop[1]           :=       0.0; // relative to rPosWait
GVL_XTS.StationParameter[nStationParameter].rReleaseDistance      :=     800.0; // relative to Mover.ActPos

nStationParameter := 76;
GVL_XTS.StationParameter[nStationParameter].eType                 := E_STATION_TYPE.STATION_PROCESS;
GVL_XTS.StationParameter[nStationParameter].sText                 := 'PROCESS_ASSEMBLY_TEST_06';
GVL_XTS.StationParameter[nStationParameter].nConfiguredStopCount  :=       1;   // how many stops the mover has to make in this station

GVL_XTS.StationParameter[nStationParameter].rPosWait              :=    21500.0+480.0; // absolute modulo position
GVL_XTS.StationParameter[nStationParameter].rPosStop[1]           :=       0.0; // relative to rPosWait
GVL_XTS.StationParameter[nStationParameter].rReleaseDistance      :=     720.0; // relative to Mover.ActPos

nStationParameter := 77;
GVL_XTS.StationParameter[nStationParameter].eType                 := E_STATION_TYPE.STATION_PROCESS;
GVL_XTS.StationParameter[nStationParameter].sText                 := 'PROCESS_ASSEMBLY_TEST_07';
GVL_XTS.StationParameter[nStationParameter].nConfiguredStopCount  :=       1;   // how many stops the mover has to make in this station

GVL_XTS.StationParameter[nStationParameter].rPosWait              :=    21500.0+560.0; // absolute modulo position
GVL_XTS.StationParameter[nStationParameter].rPosStop[1]           :=       0.0; // relative to rPosWait
GVL_XTS.StationParameter[nStationParameter].rReleaseDistance      :=     640.0; // relative to Mover.ActPos

nStationParameter := 78;
GVL_XTS.StationParameter[nStationParameter].eType                 := E_STATION_TYPE.STATION_PROCESS;
GVL_XTS.StationParameter[nStationParameter].sText                 := 'PROCESS_ASSEMBLY_TEST_08';
GVL_XTS.StationParameter[nStationParameter].nConfiguredStopCount  :=       1;   // how many stops the mover has to make in this station

GVL_XTS.StationParameter[nStationParameter].rPosWait              :=    21500.0+640.0; // absolute modulo position
GVL_XTS.StationParameter[nStationParameter].rPosStop[1]           :=       0.0; // relative to rPosWait
GVL_XTS.StationParameter[nStationParameter].rReleaseDistance      :=     560.0; // relative to Mover.ActPos

nStationParameter := 79;
GVL_XTS.StationParameter[nStationParameter].eType                 := E_STATION_TYPE.STATION_PROCESS;
GVL_XTS.StationParameter[nStationParameter].sText                 := 'PROCESS_ASSEMBLY_TEST_09';
GVL_XTS.StationParameter[nStationParameter].nConfiguredStopCount  :=       1;   // how many stops the mover has to make in this station

GVL_XTS.StationParameter[nStationParameter].rPosWait              :=    21500.0+720.0; // absolute modulo position
GVL_XTS.StationParameter[nStationParameter].rPosStop[1]           :=       0.0; // relative to rPosWait
GVL_XTS.StationParameter[nStationParameter].rReleaseDistance      :=     480.0; // relative to Mover.ActPos

nStationParameter := 80;
GVL_XTS.StationParameter[nStationParameter].eType                 := E_STATION_TYPE.STATION_PROCESS;
GVL_XTS.StationParameter[nStationParameter].sText                 := 'PROCESS_ASSEMBLY_TEST_10';
GVL_XTS.StationParameter[nStationParameter].nConfiguredStopCount  :=       1;   // how many stops the mover has to make in this station

GVL_XTS.StationParameter[nStationParameter].rPosWait              :=    21500.0+800.0; // absolute modulo position
GVL_XTS.StationParameter[nStationParameter].rPosStop[1]           :=       0.0; // relative to rPosWait
GVL_XTS.StationParameter[nStationParameter].rReleaseDistance      :=      400.0; // relative to Mover.ActPos

nStationParameter := 81;
GVL_XTS.StationParameter[nStationParameter].eType                 := E_STATION_TYPE.STATION_PROCESS;
GVL_XTS.StationParameter[nStationParameter].sText                 := 'PROCESS_ASSEMBLY_TEST_11';
GVL_XTS.StationParameter[nStationParameter].nConfiguredStopCount  :=       1;   // how many stops the mover has to make in this station

GVL_XTS.StationParameter[nStationParameter].rPosWait              :=    21500.0+880.0; // absolute modulo position
GVL_XTS.StationParameter[nStationParameter].rPosStop[1]           :=       0.0; // relative to rPosWait
GVL_XTS.StationParameter[nStationParameter].rReleaseDistance      :=      320.0; // relative to Mover.ActPos

nStationParameter := 82;
GVL_XTS.StationParameter[nStationParameter].eType                 := E_STATION_TYPE.STATION_PROCESS;
GVL_XTS.StationParameter[nStationParameter].sText                 := 'PROCESS_ASSEMBLY_TEST_12';
GVL_XTS.StationParameter[nStationParameter].nConfiguredStopCount  :=       1;   // how many stops the mover has to make in this station

GVL_XTS.StationParameter[nStationParameter].rPosWait              :=    21500.0+960.0; // absolute modulo position
GVL_XTS.StationParameter[nStationParameter].rPosStop[1]           :=       0.0; // relative to rPosWait
GVL_XTS.StationParameter[nStationParameter].rReleaseDistance      :=    240.0; // relative to Mover.ActPos

nStationParameter := 83;
GVL_XTS.StationParameter[nStationParameter].eType                 := E_STATION_TYPE.STATION_PROCESS;
GVL_XTS.StationParameter[nStationParameter].sText                 := 'PROCESS_ASSEMBLY_TEST_13';
GVL_XTS.StationParameter[nStationParameter].nConfiguredStopCount  :=       1;   // how many stops the mover has to make in this station

GVL_XTS.StationParameter[nStationParameter].rPosWait              :=    21500.0+1040.0; // absolute modulo position
GVL_XTS.StationParameter[nStationParameter].rPosStop[1]           :=       0.0; // relative to rPosWait
GVL_XTS.StationParameter[nStationParameter].rReleaseDistance      :=     160.0; // relative to Mover.ActPos

nStationParameter := 84;
GVL_XTS.StationParameter[nStationParameter].eType                 := E_STATION_TYPE.STATION_PROCESS;
GVL_XTS.StationParameter[nStationParameter].sText                 := 'PROCESS_ASSEMBLY_TEST_14';
GVL_XTS.StationParameter[nStationParameter].nConfiguredStopCount  :=       1;   // how many stops the mover has to make in this station

GVL_XTS.StationParameter[nStationParameter].rPosWait              :=    21500.0+1120.0; // absolute modulo position
GVL_XTS.StationParameter[nStationParameter].rPosStop[1]           :=       0.0; // relative to rPosWait
GVL_XTS.StationParameter[nStationParameter].rReleaseDistance      :=     80.0; // relative to Mover.ActPos

nStationParameter := 85;
GVL_XTS.StationParameter[nStationParameter].eType                 := E_STATION_TYPE.STATION_PROCESS;
GVL_XTS.StationParameter[nStationParameter].sText                 := 'PROCESS_ASSEMBLY_TEST_15';
GVL_XTS.StationParameter[nStationParameter].nConfiguredStopCount  :=       1;   // how many stops the mover has to make in this station

GVL_XTS.StationParameter[nStationParameter].rPosWait              :=    21500.0+1200.0; // absolute modulo position
GVL_XTS.StationParameter[nStationParameter].rPosStop[1]           :=       0.0; // relative to rPosWait
GVL_XTS.StationParameter[nStationParameter].rReleaseDistance      :=      25.0; // relative to Mover.ActPos

nStationParameter := 86;
GVL_XTS.StationParameter[nStationParameter].eType                 := E_STATION_TYPE.STATION_PROCESS;
GVL_XTS.StationParameter[nStationParameter].sText                 := 'PROCESS_ASSEMBLY_TEST_16';
GVL_XTS.StationParameter[nStationParameter].nConfiguredStopCount  :=       1;   // how many stops the mover has to make in this station

GVL_XTS.StationParameter[nStationParameter].rPosWait              :=    21500.0+1280.0; // absolute modulo position
GVL_XTS.StationParameter[nStationParameter].rPosStop[1]           :=       0.0; // relative to rPosWait
GVL_XTS.StationParameter[nStationParameter].rReleaseDistance      :=      -5.0; // relative to Mover.ActPos

//-----------------------------------------------------------------------------------------------------------------------------------------
// NOK handling
//-----------------------------------------------------------------------------------------------------------------------------------------
FOR nStationParameter := 91 TO 91
DO
  GVL_XTS.StationParameter[nStationParameter].rVelo               := 750.0;//MAIN_APP.rDefaultVeloMin;
END_FOR
nStationParameter := 91;
GVL_XTS.StationParameter[nStationParameter].eType                 := E_STATION_TYPE.STATION_PROCESS;
GVL_XTS.StationParameter[nStationParameter].sText                 := 'DISTRIBUTOR_CAMERA';
GVL_XTS.StationParameter[nStationParameter].nConfiguredStopCount  :=       1;   // how many stops the mover has to make in this station

GVL_XTS.StationParameter[nStationParameter].rPosWait              :=   23250.0; // absolute modulo position
GVL_XTS.StationParameter[nStationParameter].rPosStop[1]           :=       0.0; // relative to rPosWait
GVL_XTS.StationParameter[nStationParameter].rReleaseDistance      :=      -5.0; // relative to Mover.ActPos

//-----------------------------------------------------------------------------------------------------------------------------------------
// camera inspection 
//-----------------------------------------------------------------------------------------------------------------------------------------
FOR nStationParameter := 95 TO 95
DO
  GVL_XTS.StationParameter[nStationParameter].rVelo               := MAIN_APP.rDefaultVeloMin;
END_FOR
nStationParameter := 95;
GVL_XTS.StationParameter[nStationParameter].eType                 := E_STATION_TYPE.STATION_PROCESS;
GVL_XTS.StationParameter[nStationParameter].sText                 := 'CONTINUOUS_ASSEMBLY_CAMERA';
GVL_XTS.StationParameter[nStationParameter].nConfiguredStopCount  :=       1;   // how many stops the mover has to make in this station

GVL_XTS.StationParameter[nStationParameter].rPosWait              :=   24000.0+80.0; // absolute modulo position
GVL_XTS.StationParameter[nStationParameter].rPosStop[1]           :=       0.0; // relative to rPosWait
GVL_XTS.StationParameter[nStationParameter].rReleaseDistance      :=      -5.0; // relative to Mover.ActPos
GVL_XTS.StationParameter[nStationParameter].rVelo                 :=     750.0;
GVL_XTS.StationParameter[nStationParameter].rGap                  :=      78.0;

//-----------------------------------------------------------------------------------------------------------------------------------------
// DISTRIBUTOR - unloading
//-----------------------------------------------------------------------------------------------------------------------------------------
nStationParameter := 119;
GVL_XTS.StationParameter[nStationParameter].eType                 := E_STATION_TYPE.STATION_PROCESS;
GVL_XTS.StationParameter[nStationParameter].sText                 := 'DISTRIBUTOR_OUTFEED';
GVL_XTS.StationParameter[nStationParameter].nConfiguredStopCount  :=       1;   // how many stops the mover has to make in this station

GVL_XTS.StationParameter[nStationParameter].rPosWait              :=   26000.0; // absolute modulo position
GVL_XTS.StationParameter[nStationParameter].rPosStop[1]           :=       0.0; // relative to rPosWait
GVL_XTS.StationParameter[nStationParameter].rReleaseDistance      :=      -5.0; // relative to Mover.ActPos
GVL_XTS.StationParameter[nStationParameter].rVelo                 :=    1000.0;//MAIN_APP.rDefaultVeloMin;


//-----------------------------------------------------------------------------------------------------------------------------------------
// PROCESS_OUTFEED
//-----------------------------------------------------------------------------------------------------------------------------------------
FOR nStationParameter := 120 TO 133
DO
  GVL_XTS.StationParameter[nStationParameter].rVelo               := 1000.0;//MAIN_APP.rDefaultVeloMin;
END_FOR
nStationParameter := 120;
GVL_XTS.StationParameter[nStationParameter].eType                 := E_STATION_TYPE.STATION_PROCESS;
GVL_XTS.StationParameter[nStationParameter].sText                 := 'PROCESS_OUTFEED_01';
GVL_XTS.StationParameter[nStationParameter].nConfiguredStopCount  :=       1;   // how many stops the mover has to make in this station

GVL_XTS.StationParameter[nStationParameter].rPosWait              :=   26250.0; // absolute modulo position
GVL_XTS.StationParameter[nStationParameter].rPosStop[1]           :=      80.0; // relative to rPosWait
GVL_XTS.StationParameter[nStationParameter].rReleaseDistance      :=     960.0; // relative to Mover.ActPos

nStationParameter := 121;
GVL_XTS.StationParameter[nStationParameter].eType                 := E_STATION_TYPE.STATION_PROCESS;
GVL_XTS.StationParameter[nStationParameter].sText                 := 'PROCESS_OUTFEED_02';
GVL_XTS.StationParameter[nStationParameter].nConfiguredStopCount  :=       1;   // how many stops the mover has to make in this station

GVL_XTS.StationParameter[nStationParameter].rPosWait              :=   26250.0; // absolute modulo position
GVL_XTS.StationParameter[nStationParameter].rPosStop[1]           :=     160.0; // relative to rPosWait
GVL_XTS.StationParameter[nStationParameter].rReleaseDistance      :=     880.0; // relative to Mover.ActPos

nStationParameter := 122;
GVL_XTS.StationParameter[nStationParameter].eType                 := E_STATION_TYPE.STATION_PROCESS;
GVL_XTS.StationParameter[nStationParameter].sText                 := 'PROCESS_OUTFEED_03';
GVL_XTS.StationParameter[nStationParameter].nConfiguredStopCount  :=       1;   // how many stops the mover has to make in this station

GVL_XTS.StationParameter[nStationParameter].rPosWait              :=   26250.0; // absolute modulo position
GVL_XTS.StationParameter[nStationParameter].rPosStop[1]           :=     240.0; // relative to rPosWait
GVL_XTS.StationParameter[nStationParameter].rReleaseDistance      :=     800.0; // relative to Mover.ActPos

nStationParameter := 123;
GVL_XTS.StationParameter[nStationParameter].eType                 := E_STATION_TYPE.STATION_PROCESS;
GVL_XTS.StationParameter[nStationParameter].sText                 := 'PROCESS_OUTFEED_04';
GVL_XTS.StationParameter[nStationParameter].nConfiguredStopCount  :=       1;   // how many stops the mover has to make in this station

GVL_XTS.StationParameter[nStationParameter].rPosWait              :=   26250.0; // absolute modulo position
GVL_XTS.StationParameter[nStationParameter].rPosStop[1]           :=     320.0; // relative to rPosWait
GVL_XTS.StationParameter[nStationParameter].rReleaseDistance      :=     720.0; // relative to Mover.ActPos

nStationParameter := 124;
GVL_XTS.StationParameter[nStationParameter].eType                 := E_STATION_TYPE.STATION_PROCESS;
GVL_XTS.StationParameter[nStationParameter].sText                 := 'PROCESS_OUTFEED_05';
GVL_XTS.StationParameter[nStationParameter].nConfiguredStopCount  :=       1;   // how many stops the mover has to make in this station

GVL_XTS.StationParameter[nStationParameter].rPosWait              :=   26250.0; // absolute modulo position
GVL_XTS.StationParameter[nStationParameter].rPosStop[1]           :=     400.0; // relative to rPosWait
GVL_XTS.StationParameter[nStationParameter].rReleaseDistance      :=     640.0; // relative to Mover.ActPos

nStationParameter := 125;
GVL_XTS.StationParameter[nStationParameter].eType                 := E_STATION_TYPE.STATION_PROCESS;
GVL_XTS.StationParameter[nStationParameter].sText                 := 'PROCESS_OUTFEED_06';
GVL_XTS.StationParameter[nStationParameter].nConfiguredStopCount  :=       1;   // how many stops the mover has to make in this station

GVL_XTS.StationParameter[nStationParameter].rPosWait              :=   26250.0; // absolute modulo position
GVL_XTS.StationParameter[nStationParameter].rPosStop[1]           :=     480.0; // relative to rPosWait
GVL_XTS.StationParameter[nStationParameter].rReleaseDistance      :=     560.0; // relative to Mover.ActPos

nStationParameter := 126;
GVL_XTS.StationParameter[nStationParameter].eType                 := E_STATION_TYPE.STATION_PROCESS;
GVL_XTS.StationParameter[nStationParameter].sText                 := 'PROCESS_OUTFEED_07';
GVL_XTS.StationParameter[nStationParameter].nConfiguredStopCount  :=       1;   // how many stops the mover has to make in this station

GVL_XTS.StationParameter[nStationParameter].rPosWait              :=   26250.0; // absolute modulo position
GVL_XTS.StationParameter[nStationParameter].rPosStop[1]           :=     560.0; // relative to rPosWait
GVL_XTS.StationParameter[nStationParameter].rReleaseDistance      :=     480.0; // relative to Mover.ActPos

nStationParameter := 127;
GVL_XTS.StationParameter[nStationParameter].eType                 := E_STATION_TYPE.STATION_PROCESS;
GVL_XTS.StationParameter[nStationParameter].sText                 := 'PROCESS_OUTFEED_08';
GVL_XTS.StationParameter[nStationParameter].nConfiguredStopCount  :=       1;   // how many stops the mover has to make in this station

GVL_XTS.StationParameter[nStationParameter].rPosWait              :=   26250.0; // absolute modulo position
GVL_XTS.StationParameter[nStationParameter].rPosStop[1]           :=     640.0; // relative to rPosWait
GVL_XTS.StationParameter[nStationParameter].rReleaseDistance      :=     400.0; // relative to Mover.ActPos

nStationParameter := 128;
GVL_XTS.StationParameter[nStationParameter].eType                 := E_STATION_TYPE.STATION_PROCESS;
GVL_XTS.StationParameter[nStationParameter].sText                 := 'PROCESS_OUTFEED_09';
GVL_XTS.StationParameter[nStationParameter].nConfiguredStopCount  :=       1;   // how many stops the mover has to make in this station

GVL_XTS.StationParameter[nStationParameter].rPosWait              :=   26250.0; // absolute modulo position
GVL_XTS.StationParameter[nStationParameter].rPosStop[1]           :=     720.0; // relative to rPosWait
GVL_XTS.StationParameter[nStationParameter].rReleaseDistance      :=     320.0; // relative to Mover.ActPos

nStationParameter := 129;
GVL_XTS.StationParameter[nStationParameter].eType                 := E_STATION_TYPE.STATION_PROCESS;
GVL_XTS.StationParameter[nStationParameter].sText                 := 'PROCESS_OUTFEED_10';
GVL_XTS.StationParameter[nStationParameter].nConfiguredStopCount  :=       1;   // how many stops the mover has to make in this station

GVL_XTS.StationParameter[nStationParameter].rPosWait              :=   26250.0; // absolute modulo position
GVL_XTS.StationParameter[nStationParameter].rPosStop[1]           :=     800.0; // relative to rPosWait
GVL_XTS.StationParameter[nStationParameter].rReleaseDistance      :=     240.0; // relative to Mover.ActPos

nStationParameter := 130;
GVL_XTS.StationParameter[nStationParameter].eType                 := E_STATION_TYPE.STATION_PROCESS;
GVL_XTS.StationParameter[nStationParameter].sText                 := 'PROCESS_OUTFEED_11';
GVL_XTS.StationParameter[nStationParameter].nConfiguredStopCount  :=       1;   // how many stops the mover has to make in this station

GVL_XTS.StationParameter[nStationParameter].rPosWait              :=   26250.0; // absolute modulo position
GVL_XTS.StationParameter[nStationParameter].rPosStop[1]           :=     880.0; // relative to rPosWait
GVL_XTS.StationParameter[nStationParameter].rReleaseDistance      :=     160.0; // relative to Mover.ActPos

nStationParameter := 131;
GVL_XTS.StationParameter[nStationParameter].eType                 := E_STATION_TYPE.STATION_PROCESS;
GVL_XTS.StationParameter[nStationParameter].sText                 := 'PROCESS_OUTFEED_12';
GVL_XTS.StationParameter[nStationParameter].nConfiguredStopCount  :=       1;   // how many stops the mover has to make in this station

GVL_XTS.StationParameter[nStationParameter].rPosWait              :=   26250.0; // absolute modulo position
GVL_XTS.StationParameter[nStationParameter].rPosStop[1]           :=     960.0; // relative to rPosWait
GVL_XTS.StationParameter[nStationParameter].rReleaseDistance      :=     80.0; // relative to Mover.ActPos

nStationParameter := 132;
GVL_XTS.StationParameter[nStationParameter].eType                 := E_STATION_TYPE.STATION_PROCESS;
GVL_XTS.StationParameter[nStationParameter].sText                 := 'PROCESS_OUTFEED_13';
GVL_XTS.StationParameter[nStationParameter].nConfiguredStopCount  :=       1;   // how many stops the mover has to make in this station

GVL_XTS.StationParameter[nStationParameter].rPosWait              :=   26250.0; // absolute modulo position
GVL_XTS.StationParameter[nStationParameter].rPosStop[1]           :=    1040.0; // relative to rPosWait
GVL_XTS.StationParameter[nStationParameter].rReleaseDistance      :=      25.0; // relative to Mover.ActPos

nStationParameter := 133;
GVL_XTS.StationParameter[nStationParameter].eType                 := E_STATION_TYPE.STATION_PROCESS;
GVL_XTS.StationParameter[nStationParameter].sText                 := 'PROCESS_OUTFEED_14';
GVL_XTS.StationParameter[nStationParameter].nConfiguredStopCount  :=       1;   // how many stops the mover has to make in this station

GVL_XTS.StationParameter[nStationParameter].rPosWait              :=   26250.0; // absolute modulo position
GVL_XTS.StationParameter[nStationParameter].rPosStop[1]           :=    1120.0; // relative to rPosWait
GVL_XTS.StationParameter[nStationParameter].rReleaseDistance      :=      -5.0; // relative to Mover.ActPos

//-----------------------------------------------------------------------------------------------------------------------------------------
//  DISTRIBUTOR
//-----------------------------------------------------------------------------------------------------------------------------------------
nStationParameter := 140;
GVL_XTS.StationParameter[nStationParameter].eType                 := E_STATION_TYPE.STATION_PROCESS;
GVL_XTS.StationParameter[nStationParameter].sText                 := 'DISTRIBUTOR_WPC_CLEAN';
GVL_XTS.StationParameter[nStationParameter].nConfiguredStopCount  :=      1;   // how many stops the mover has to make in this station

GVL_XTS.StationParameter[nStationParameter].rPosWait              :=   1000.0; // absolute modulo position
GVL_XTS.StationParameter[nStationParameter].rPosStop[1]           :=      0.0; // relative to rPosWait
GVL_XTS.StationParameter[nStationParameter].rReleaseDistance      :=     -5.0; // relative to Mover.ActPos

GVL_XTS.StationParameter[nStationParameter].rGap                  :=    100.0;
GVL_XTS.StationParameter[nStationParameter].rVelo                 :=   2500.0;
GVL_XTS.StationParameter[nStationParameter].rAccDec               :=  17500.0;
GVL_XTS.StationParameter[nStationParameter].rJerk                 :=  300000.0;

//-----------------------------------------------------------------------------------------------------------------------------------------
//  PRC 14 wpc clean
//-----------------------------------------------------------------------------------------------------------------------------------------
nStationParameter := 141;
GVL_XTS.StationParameter[nStationParameter].eType                 := E_STATION_TYPE.STATION_PROCESS;
GVL_XTS.StationParameter[nStationParameter].sText                 := 'CONTINUOUS_WPC_CLEAN';
GVL_XTS.StationParameter[nStationParameter].nConfiguredStopCount  :=      1;   // how many stops the mover has to make in this station

GVL_XTS.StationParameter[nStationParameter].rPosWait              :=   4000.0; // absolute modulo position
GVL_XTS.StationParameter[nStationParameter].rPosStop[1]           :=      0.0; // relative to rPosWait
GVL_XTS.StationParameter[nStationParameter].rReleaseDistance      :=      -5.0; // relative to Mover.ActPos
GVL_XTS.StationParameter[nStationParameter].rVelo                 :=     750.0;
GVL_XTS.StationParameter[nStationParameter].rGap                  :=     100.0;
GVL_XTS.StationParameter[nStationParameter].rJerk                 :=  300000.0;

//-----------------------------------------------------------------------------------------------------------------------------------------
//  DISTRIBUTOR
//-----------------------------------------------------------------------------------------------------------------------------------------
nStationParameter := 142;
GVL_XTS.StationParameter[nStationParameter].eType                 := E_STATION_TYPE.STATION_PROCESS;
GVL_XTS.StationParameter[nStationParameter].sText                 := 'DISTRIBUTOR_INFEED';
GVL_XTS.StationParameter[nStationParameter].nConfiguredStopCount  :=      1;   // how many stops the mover has to make in this station

GVL_XTS.StationParameter[nStationParameter].rPosWait              :=   5500.0; // absolute modulo position
GVL_XTS.StationParameter[nStationParameter].rPosStop[1]           :=      0.0; // relative to rPosWait
GVL_XTS.StationParameter[nStationParameter].rReleaseDistance      :=    -10.0; // relative to Mover.ActPos

GVL_XTS.StationParameter[nStationParameter].rGap                  :=     78.0;
GVL_XTS.StationParameter[nStationParameter].rVelo                 :=   1500.0;

//-----------------------------------------------------------------------------------------------------------------------------------------
//-----------------------------------------------------------------------------------------------------------------------------------------
// EOF
//-----------------------------------------------------------------------------------------------------------------------------------------
//-----------------------------------------------------------------------------------------------------------------------------------------

END_FUNCTION

(* stored: Version 1.1.0.1, ProductVersion 3.1.4026.20
   POU StationParameter_28000_1: Id {066966a3-913e-4d6a-a6dc-2f2d207e3fa2}, SpecialFunc None *)
